Fanuc KAREL source: KC00002.KL

PROGRAM KC00002
%NOLOCKGROUP
%ENVIRONMENT PC
VAR
  I: INTEGER
  J: INTEGER
  K: INTEGER
  R: REAL
  B: BOOLEAN
  S: STRING[80]
  T: STRING[80]
  P: PATH
  Q: PATH
  AI: ARRAY[8] OF INTEGER
  AB: ARRAY[244] OF BYTE
BEGIN
  ADD_INTPC(AB,I,J,K)
END KC00002
